(* IEC 61131-3 sources: plc-iiot-stack/src/POUs/Iiot/F_IiotDeadbandExceeded, 2 files *)

(* ---- F_IiotDeadbandExceeded.decl.st ---- *)
// Назначение: значение ушло от последнего опубликованного больше зоны нечувствительности:
//             |новое - последнее| > зона (строго больше; зона <= 0 или не число — любое изменение).
//             Переход между конечным и неконечным значением — изменение, два неконечных — нет.
// Автор:      kr0nsch
// Версия:     0.1.0
// Документ:   docs/plc_mqtt.md, раздел «Телеметрия»
FUNCTION F_IiotDeadbandExceeded : BOOL
VAR_INPUT
    lrNew : LREAL;      // текущее значение
    lrLast : LREAL;     // последнее опубликованное
    rDeadband : REAL;   // зона нечувствительности, в единицах значения
END_VAR
VAR
    xNewFinite : BOOL;
    xLastFinite : BOOL;
    lrDiff : LREAL;
END_VAR

(* ---- F_IiotDeadbandExceeded.impl.st ---- *)
xNewFinite := F_IsFiniteLreal(lrValue := lrNew);
xLastFinite := F_IsFiniteLreal(lrValue := lrLast);
IF NOT xNewFinite OR NOT xLastFinite THEN
    F_IiotDeadbandExceeded := xNewFinite <> xLastFinite;
    RETURN;
END_IF
lrDiff := ABS(lrNew - lrLast);
IF NOT F_IsFiniteReal(rValue := rDeadband) OR rDeadband <= 0.0 THEN
    F_IiotDeadbandExceeded := lrDiff > 0.0;
ELSE
    F_IiotDeadbandExceeded := lrDiff > REAL_TO_LREAL(rDeadband);
END_IF
